Fanuc KAREL source: ko00051.KL

-- PROVISIONAL review KL for V1013-1; original PC SHA256 1b3efa3cce46ac592ccc9c92e60181d754d90072c6bf14ef60d7484271320ddb
-- Incomplete behavior may be omitted. Consult companion uncertainty JSON. Do not deploy.
PROGRAM KO00051
%NOLOCKGROUP
BEGIN
  -- UNRESOLVED_PC offsets 5-12; opcodes 9D,23
  -- UNRESOLVED_PC offsets 17-66; opcodes 27,27,49,7E,AD,22,1C,22,31,7E,4A
  -- UNRESOLVED_PC offsets 71-75; opcodes 7F
END KO00051
